TYPE ST_Road :
STRUCT
	nId: UINT;
	fLength: LREAL;
END_STRUCT
END_TYPE

(* stored: Version 1.1.0.1, ProductVersion 3.1.4024.12
   DUT ST_Road: Id {bfcdb122-ad7e-4a01-afc7-4015e7d44e02} *)
